(* IEC 61131-3 sources: volt/packages/volt-lsp-iec/test-corpus/twincat-project14/TwinCAT Project14/PLC/Untitled2/Untitled2 Project/POUs, 4 files *)

(* ---- VltFixtureCfc.pou ---- *)
FUNCTION_BLOCK VltFixtureCfc
VAR_INPUT
END_VAR
VAR_OUTPUT
END_VAR
VAR
END_VAR
%LANGUAGE CFC UNSUPPORTED

END_FUNCTION_BLOCK

(* ---- VltFixtureMembers.pou ---- *)
FUNCTION_BLOCK VltFixtureMembers
VAR_INPUT
	bGo : BOOL;
END_VAR
VAR
	nTick : INT;
END_VAR

%LANGUAGE ST
nTick := nTick + 1;

END_FUNCTION_BLOCK

METHOD CfcStep : BOOL
VAR_INPUT
	bIn : BOOL;
END_VAR

%LANGUAGE CFC UNSUPPORTED
END_METHOD

METHOD Visible : BOOL
VAR_INPUT
	bIn : BOOL;
END_VAR

%LANGUAGE ST
Visible := bIn;
END_METHOD

ACTION SfcRun
%LANGUAGE SFC UNSUPPORTED
END_ACTION

(* ---- VltFixtureSfc.pou ---- *)
FUNCTION_BLOCK VltFixtureSfc
VAR_INPUT
END_VAR
VAR_OUTPUT
END_VAR
VAR
END_VAR
%LANGUAGE SFC UNSUPPORTED

END_FUNCTION_BLOCK

(* ---- POUexecute.pou ---- *)
PROGRAM POUexecute
VAR
	iCount:INT;

	t1: TON;
	output: BOOL;
	e1: TIME;
	in1: BOOL;
	a: BOOL;
	b: BOOL;
	c: BOOL;
	out1: BOOL;
	t2: TON;
	out2: INT;
END_VAR
%LANGUAGE LD
%NETWORK
EXECUTE(EN := TRUE, 'iCount:=icount+1;
');
%NETWORK
ASSIGN(t1(IN := in1, PT := e1), Q => output);
%NETWORK
VAR w1 : ANY; END_VAR
w1 := b;
ASSIGN(AND(OR(a, w1), c), Q => out1);
ASSIGN(w1, Q => out2);
%NETWORK
ASSIGN(t2(PT := e1), Q => output);

END_PROGRAM
